{attribute 'qualified_only'}
{attribute 'strict'}
TYPE E_ConveyorMode  :
(
	AUTO,
	MANUAL
);
END_TYPE

(* stored: Version 1.1.0.1, ProductVersion 3.1.4024.16
   DUT E_ConveyorMode: Id {773c6bf0-794b-44ea-86e7-65b49d22e565} *)
